// TIA Portal V19 export
FUNCTION_BLOCK "Sim_SMOutputs"   // FB6, FBD
{ S7_Optimized_Access := 'TRUE' }
// stored: MemoryReserve 100, SetENOAutomatically false
   VAR
      VaccumPID { ExternalAccessible := 'False'; ExternalVisible := 'False'; ExternalWritable := 'False'} : "PidL";
      SteamPID { S7_SetPoint := 'True'} : "PidL";
      SimularDelay { S7_SetPoint := 'True'} : TON_TIME;
      FeedPID { S7_SetPoint := 'True'} : "PidL";
      LiSet : Bool;
      LiSetM : Bool;
      LevelInit : Real;
      BrixInit : Real;
   END_VAR
   // VaccumPID.AutModLi := true;
   // VaccumPID.ModLiOp := true;
   // VaccumPID.PV_Norm.High := 2000.0;
   // VaccumPID.PV_Scale.High := 2000.0;
   // VaccumPID.DataHMI.SpInt := 200.0;
   // VaccumPID.DataHMI.PIDConfig.NegGain := true;
   // VaccumPID.DataHMI.PIDConfig.Ti := 80.0;
   // VaccumPID.DataHMI.PIDConfig.Td := 0.0;
   // VaccumPID.DataHMI.PIDConfig.DeadBW := 5.0;
   // SteamPID.AutModLi := true;
   // SteamPID.ModLiOp := true;
   // SteamPID.SPModLiOp := true;
   // SteamPID.ExtModLi := true;
   // SteamPID.SPExt := 80.0;
   // SteamPID.DataHMI.PIDConfig.Ti := 80.0;
   // FeedPID.AutModLi := true;
   // FeedPID.ModLiOp := true;
   VAR_TEMP   // added for the SCL form of the ladder/FBD networks
      _w1 : Bool;
   END_VAR
BEGIN

REGION Network 1: delay
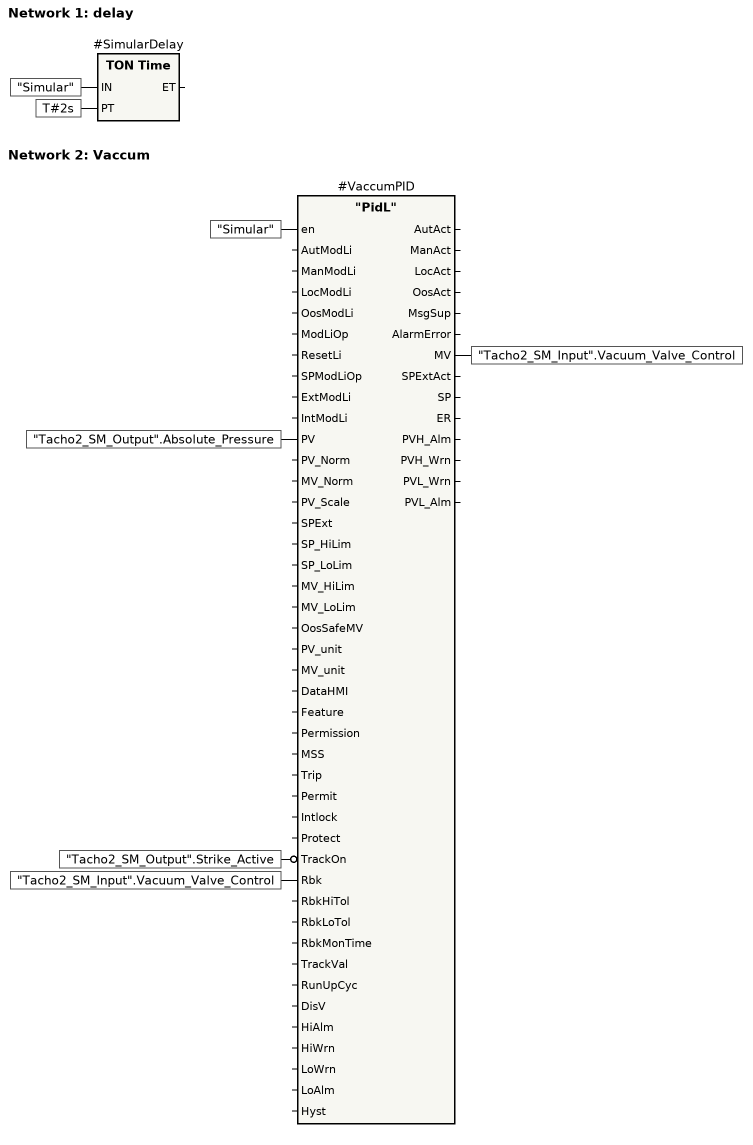
   #SimularDelay(IN := "Simular", PT := T#2s);   // TON
END_REGION

REGION Network 2: Vaccum
   IF "Simular" THEN
       #VaccumPID(PV := "Tacho2_SM_Output".Absolute_Pressure,   // "PidL"
                  TrackOn := NOT "Tacho2_SM_Output".Strike_Active,
                  Rbk := "Tacho2_SM_Input".Vacuum_Valve_Control,
                  MV => "Tacho2_SM_Input".Vacuum_Valve_Control);
   END_IF;
END_REGION

REGION Network 3: Steam
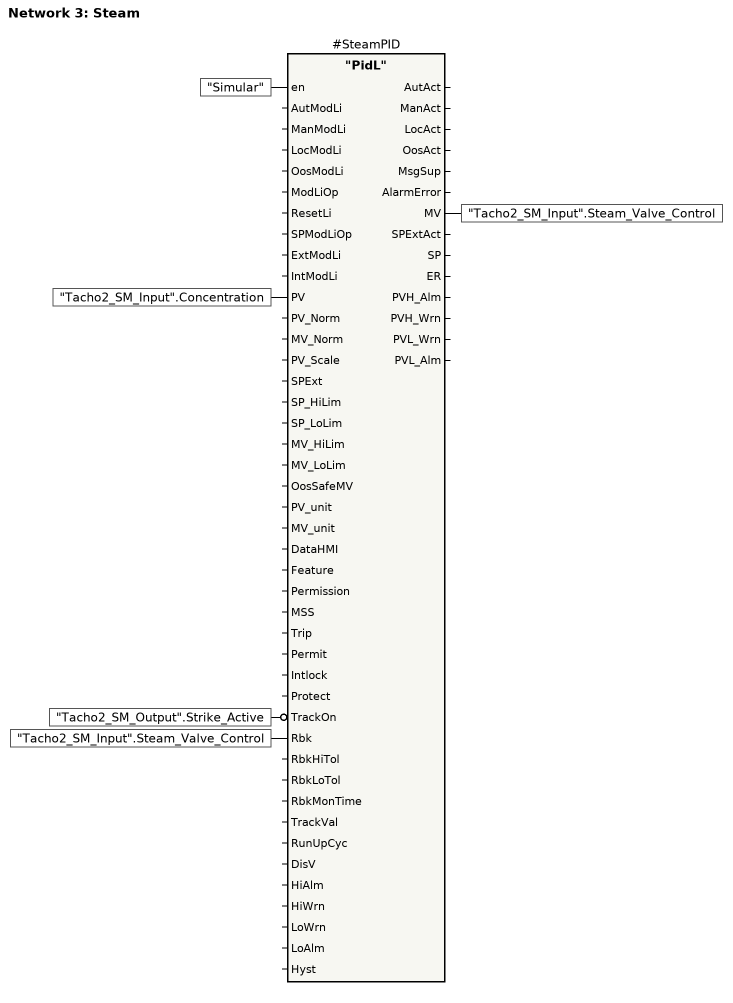
   IF "Simular" THEN
       #SteamPID(PV := "Tacho2_SM_Input".Concentration,   // "PidL"
                 TrackOn := NOT "Tacho2_SM_Output".Strike_Active,
                 Rbk := "Tacho2_SM_Input".Steam_Valve_Control,
                 MV => "Tacho2_SM_Input".Steam_Valve_Control);
   END_IF;
END_REGION

REGION Network 4
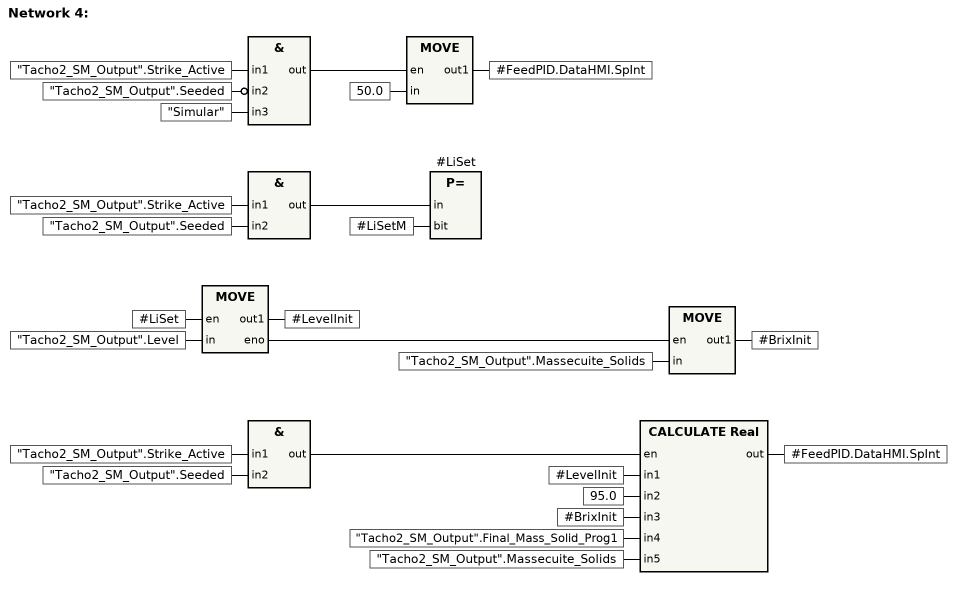
   IF "Tacho2_SM_Output".Strike_Active AND NOT "Tacho2_SM_Output".Seeded AND "Simular" THEN
       #FeedPID.DataHMI.SpInt := 50.0;
   END_IF;
   #_w1 := "Tacho2_SM_Output".Strike_Active AND "Tacho2_SM_Output".Seeded;
   #LiSet := #_w1 AND NOT #LiSetM;   // rising edge
   #LiSetM := #_w1;
   IF #LiSet THEN
       #LevelInit := "Tacho2_SM_Output".Level;
       #BrixInit := "Tacho2_SM_Output".Massecuite_Solids;
   END_IF;
   IF "Tacho2_SM_Output".Strike_Active AND "Tacho2_SM_Output".Seeded THEN
       #FeedPID.DataHMI.SpInt := #LevelInit + ((95.0 - #LevelInit)*(("Tacho2_SM_Output".Massecuite_Solids-#BrixInit)/("Tacho2_SM_Output".Final_Mass_Solid_Prog1-#BrixInit)));
   END_IF;
END_REGION

REGION Network 5
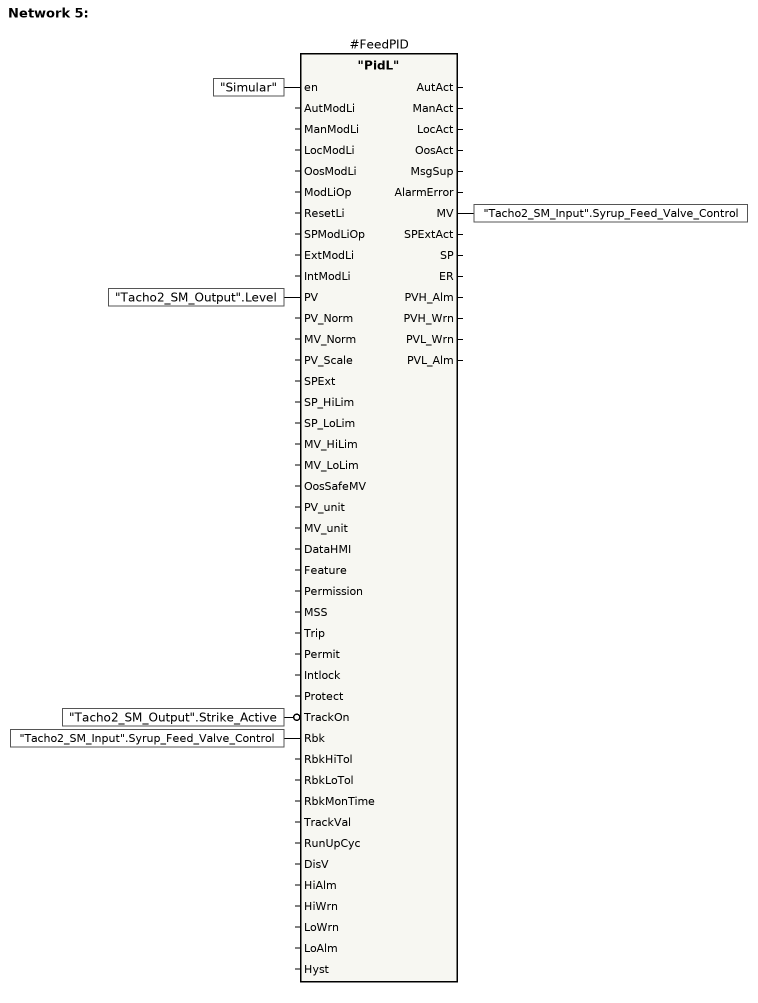
   IF "Simular" THEN
       #FeedPID(PV := "Tacho2_SM_Output".Level,   // "PidL"
                TrackOn := NOT "Tacho2_SM_Output".Strike_Active,
                Rbk := "Tacho2_SM_Input".Syrup_Feed_Valve_Control,
                MV => "Tacho2_SM_Input".Syrup_Feed_Valve_Control);
   END_IF;
END_REGION
END_FUNCTION_BLOCK
